(* Logix 5000 project; controller DSFW_0512_C_FCB_S1_SPN vendor 1 type 14 code 77 rev 20.12; software revision 20.06; part 2 of 3 *)
(* tags used below, declared in another part *)
   Alarms : DINT[3];
   Batch_Mode_Enable : BOOL;
   Comp_Low_Pressure_Alarm_Setpoint : REAL;
   Compressor_High_Pressure_Alarm_Setpoint : REAL;
   Compressor_High_Pressure_Delay_Timer : TIMER;
   Compressor_High_Superheat_Alarm_Delay : TIMER;
   Compressor_High_Superheat_Alarm_Setpoint : REAL;
   Compressor_Low_Pressure_Delay_Timer : TIMER;
   Compressor_Low_Subcooling_Alarm_Delay : TIMER;
   Compressor_Low_Subcooling_Alarm_Setpoint : REAL;
   Compressor_Low_Superheat_Alarm_Delay : TIMER;
   Compressor_Low_Superheat_Alarm_Setpoint : REAL;
   Compressor_OK_To_Run : BOOL;
   Compressor_Run_Proof_Delay : TIMER;
   Compressor_Short_Cycle_Time_Remaining : REAL;
   Compressor_Short_Cycle_Timer : TIMER;
   Compressor_Start_Delay : TIMER;
   Compressor_Subcooling : REAL;
   Compressor_Superheat : REAL;
   DV_IN_N7_100_199 : INT[10];
   DV_OUT_N7_0_99 : INT[20];
   EEV_101_Pressure_PIDE : PID_ENHANCED;
   EEV_101_Range_1_Max : REAL;
   EEV_101_Range_1_Min : REAL;
   EEV_101_Range_2_Max : REAL;
   EEV_101_Range_2_Min : REAL;
   EEV_101_Range_3_Max : REAL;
   EEV_101_Range_3_Min : REAL;
   EEV_101_Run_PIDE : BOOL;
   EEV_101_Run_Temp_PIDE : BOOL;
   EEV_101_Stop_PIDE : BOOL;
   EEV_101_Superheat_PIDE : PID_ENHANCED;
   EEV_101_Temperature_PIDE : PID_ENHANCED;
   EEV_102_Stop_PIDE : BOOL;
   Enable_Batch : BOOL;
   Evaporator_Superheat : REAL;
   Heaters_OK_To_Run : BOOL;
   Large_Batch_Derivative : REAL;
   Large_Batch_Integral : REAL;
   Large_Batch_Proportional : REAL;
   Large_Batch_Selected : BOOL;
   Medium_Batch_Derivative : REAL;
   Medium_Batch_Integral : REAL;
   Medium_Batch_Proportional : REAL;
   Medium_Batch_Selected : BOOL;
   PT_101_Offset : REAL;
   PT_101_Reactor_Supply_Pressure : REAL;
   PT_102_Compressor_Suction_Pressure : REAL;
   PT_102_Sensor_Alarm_Delay : TIMER;
   PT_103_Compressor_Discharge_Pressure : REAL;
   PT_103_Sensor_Alarm_Delay : TIMER;
   PT_104_Evaporator_Suction_Pressure : REAL;
   PT_104_Sensor_Alarm_Delay : TIMER;
   PT_105_Offset : REAL;
   PT_105_Tank_Blanket_Pressure : REAL;
   Pump_OK_To_Run : BOOL;
   Reaactor_Batch_PIDE : PID_ENHANCED;
   Reactor_Batch_CV_as_SP : REAL;
   Reactor_Batch_PID_Start : BOOL;
   Reactor_Batch_PID_Start_Delay : TIMER;
   Reactor_Batch_PID_Start_ONS : BOOL;
   Reactor_Batch_PID_Stop : BOOL;
   Reactor_Batch_PV : REAL;
   Reactor_Batch_SP_High : REAL;
   Reactor_Batch_SP_Low : REAL;
   Remote_Enable : BOOL;
   Remote_Start : BOOL;
   SCR_101_Auto_Manual : BOOL;
   SCR_101_Manual_Output : REAL;
   SCR_101_Run_PIDE : BOOL;
   SCR_101_Stop_PIDE : BOOL;
   SIC_101_Auto_Manual : BOOL;
   SIC_101_Manual_Output : REAL;
   SIC_101_Pressure_Setpoint : REAL;
   SIC_101_Run_PIDE : BOOL;
   SIC_101_Stop_PIDE : BOOL;
   Small_Batch_Derivative : REAL;
   Small_Batch_Integral : REAL;
   Small_Batch_Proportional : REAL;
   Small_Batch_Selected : BOOL;
   SP_Add_Max : REAL;
   System_Start : BOOL;
   TCV_101_Define_Range_1_Max : REAL;
   TCV_101_Define_Range_1_Min : REAL;
   TCV_101_Define_Range_2_Max : REAL;
   TCV_101_Define_Range_2_Min : REAL;
   TCV_101_Define_Range_3_Max : REAL;
   TCV_101_Define_Range_3_Min : REAL;
   TCV_101_PIDE : PID_ENHANCED;
   TCV_101_Range_1_Max : REAL;
   TCV_101_Range_1_Min : REAL;
   TCV_101_Range_2_Max : REAL;
   TCV_101_Range_2_Min : REAL;
   TCV_101_Range_3_Max : REAL;
   TCV_101_Range_3_Min : REAL;
   TCV_101_Run_PIDE : BOOL;
   TCV_101_Stop_PIDE : BOOL;
   TE_101_Liquid_Line_Temperature : REAL;
   TE_102_Evaporator_Suction_Temperature : REAL;
   TE_103_Compressor_Suction_Temperature : REAL;
   TE_104_Offset : REAL;
   TE_104_Reactor_Return_Temperature : REAL;
   TE_105_Offset : REAL;
   TE_105_Reactor_Supply_Temperature : REAL;
   Temperature_Setpoint : REAL;
   Test_Bit : BOOL[32];
   TIT_101_Offset : REAL;
   TIT_101_Vessel_Temperature : REAL;
   TIT_201_Vessel_Temperature : REAL;
   TIT_301_Vessel_Temperature : REAL;
   Vessel_1_Scale_Max : REAL;
   Vessel_1_Scale_Min : REAL;
   Vessel_1_Selected : BOOL;
   Vessel_2_Scale_Max : REAL;
   Vessel_2_Scale_Min : REAL;
   Vessel_2_Selected : BOOL;
   Vessel_3_Scale_Max : REAL;
   Vessel_3_Scale_Min : REAL;
   Vessel_3_Selected : BOOL;
(* Process_Control, continued *)

ROUTINE Heaters_Batch_Control   (* ladder *)
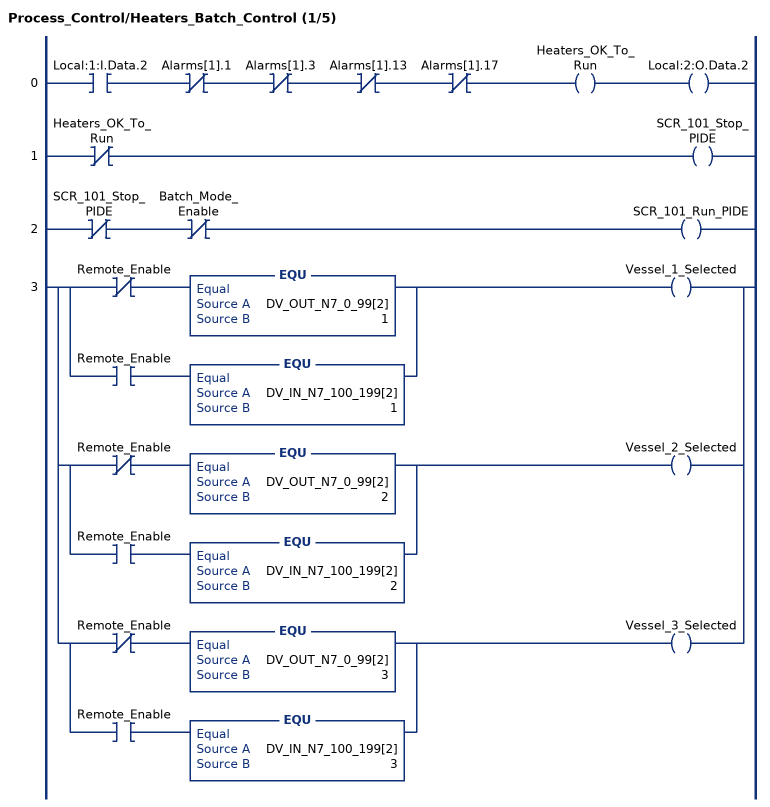
   0: XIC(Local:1:I.Data.2)XIO(Alarms[1].1)XIO(Alarms[1].3)XIO(Alarms[1].13)XIO(Alarms[1].17)OTE(Heaters_OK_To_Run)OTE(Local:2:O.Data.2);
   1: XIO(Heaters_OK_To_Run)OTE(SCR_101_Stop_PIDE);
   2: XIO(SCR_101_Stop_PIDE)XIO(Batch_Mode_Enable)OTE(SCR_101_Run_PIDE);
   3: [[XIO(Remote_Enable) EQU(DV_OUT_N7_0_99[2],1) ,XIC(Remote_Enable) EQU(DV_IN_N7_100_199[2],1) ] OTE(Vessel_1_Selected) ,[XIO(Remote_Enable) EQU(DV_OUT_N7_0_99[2],2) ,XIC(Remote_Enable) EQU(DV_IN_N7_100_199[2],2) ] OTE(Vessel_2_Selected) ,[XIO(Remote_Enable) EQU(DV_OUT_N7_0_99[2],3) ,XIC(Remote_Enable) EQU(DV_IN_N7_100_199[2],3) ] OTE(Vessel_3_Selected) ];
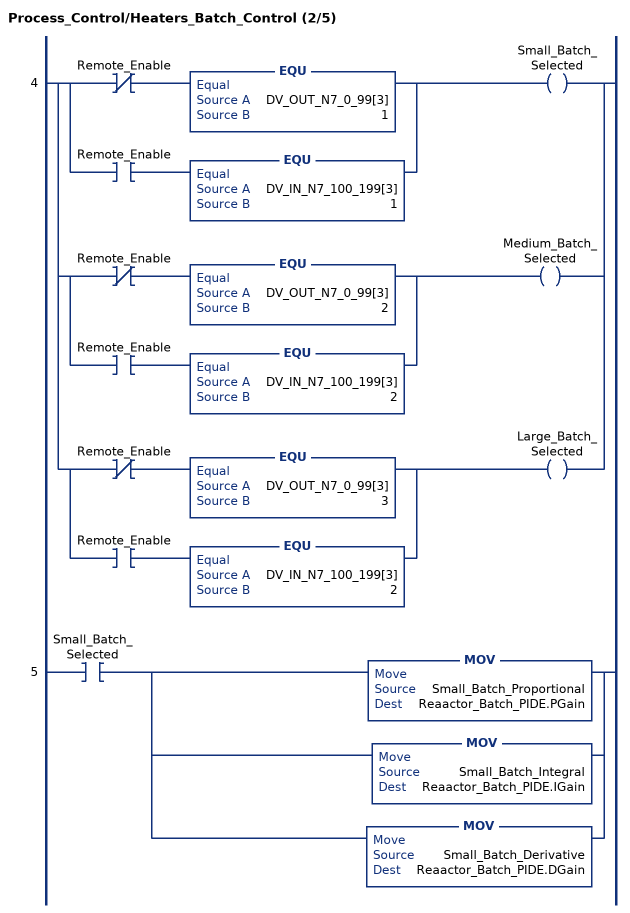
   4: [[XIO(Remote_Enable) EQU(DV_OUT_N7_0_99[3],1) ,XIC(Remote_Enable) EQU(DV_IN_N7_100_199[3],1) ] OTE(Small_Batch_Selected) ,[XIO(Remote_Enable) EQU(DV_OUT_N7_0_99[3],2) ,XIC(Remote_Enable) EQU(DV_IN_N7_100_199[3],2) ] OTE(Medium_Batch_Selected) ,[XIO(Remote_Enable) EQU(DV_OUT_N7_0_99[3],3) ,XIC(Remote_Enable) EQU(DV_IN_N7_100_199[3],2) ] OTE(Large_Batch_Selected) ];
   5: XIC(Small_Batch_Selected)[MOV(Small_Batch_Proportional,Reaactor_Batch_PIDE.PGain) ,MOV(Small_Batch_Integral,Reaactor_Batch_PIDE.IGain) ,MOV(Small_Batch_Derivative,Reaactor_Batch_PIDE.DGain) ];
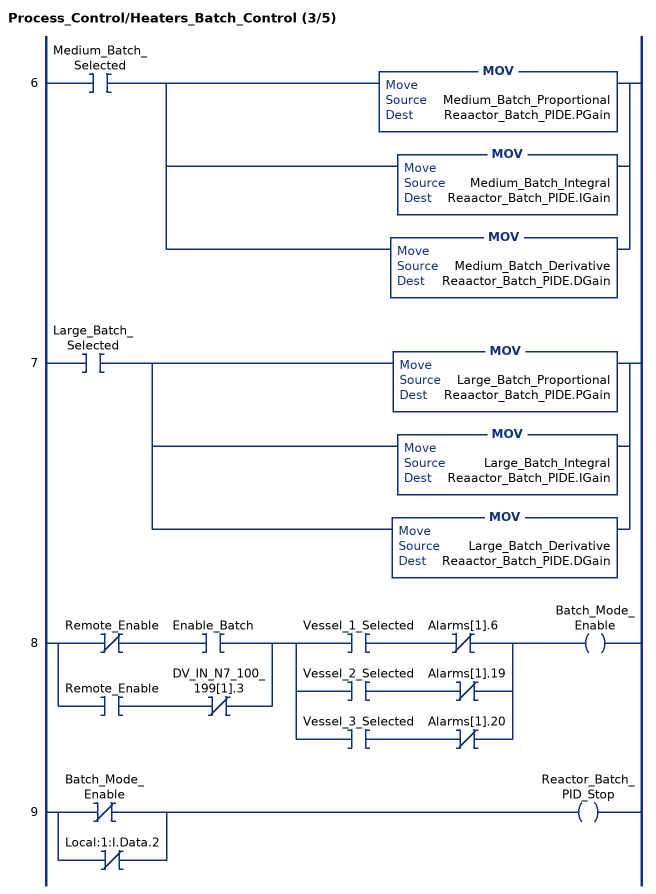
   6: XIC(Medium_Batch_Selected)[MOV(Medium_Batch_Proportional,Reaactor_Batch_PIDE.PGain) ,MOV(Medium_Batch_Integral,Reaactor_Batch_PIDE.IGain) ,MOV(Medium_Batch_Derivative,Reaactor_Batch_PIDE.DGain) ];
   7: XIC(Large_Batch_Selected)[MOV(Large_Batch_Proportional,Reaactor_Batch_PIDE.PGain) ,MOV(Large_Batch_Integral,Reaactor_Batch_PIDE.IGain) ,MOV(Large_Batch_Derivative,Reaactor_Batch_PIDE.DGain) ];
   8: [XIO(Remote_Enable) XIC(Enable_Batch) ,XIC(Remote_Enable) XIO(DV_IN_N7_100_199[1].3) ][XIC(Vessel_1_Selected) XIO(Alarms[1].6) ,XIC(Vessel_2_Selected) XIO(Alarms[1].19) ,XIC(Vessel_3_Selected) XIO(Alarms[1].20) ]OTE(Batch_Mode_Enable);
   9: [XIO(Batch_Mode_Enable) ,XIO(Local:1:I.Data.2) ]OTE(Reactor_Batch_PID_Stop);
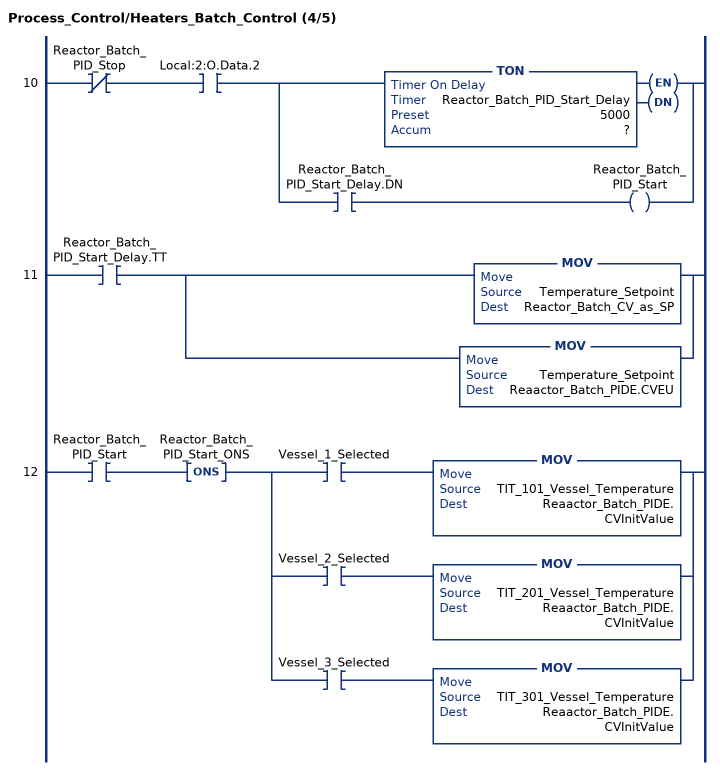
   10: XIO(Reactor_Batch_PID_Stop)XIC(Local:2:O.Data.2)[TON(Reactor_Batch_PID_Start_Delay,?,?) ,XIC(Reactor_Batch_PID_Start_Delay.DN) OTE(Reactor_Batch_PID_Start) ];
   11: XIC(Reactor_Batch_PID_Start_Delay.TT)[MOV(Temperature_Setpoint,Reactor_Batch_CV_as_SP) ,MOV(Temperature_Setpoint,Reaactor_Batch_PIDE.CVEU) ];
   12: XIC(Reactor_Batch_PID_Start)ONS(Reactor_Batch_PID_Start_ONS)[XIC(Vessel_1_Selected) MOV(TIT_101_Vessel_Temperature,Reaactor_Batch_PIDE.CVInitValue) ,XIC(Vessel_2_Selected) MOV(TIT_201_Vessel_Temperature,Reaactor_Batch_PIDE.CVInitValue) ,XIC(Vessel_3_Selected) MOV(TIT_301_Vessel_Temperature,Reaactor_Batch_PIDE.CVInitValue) ];
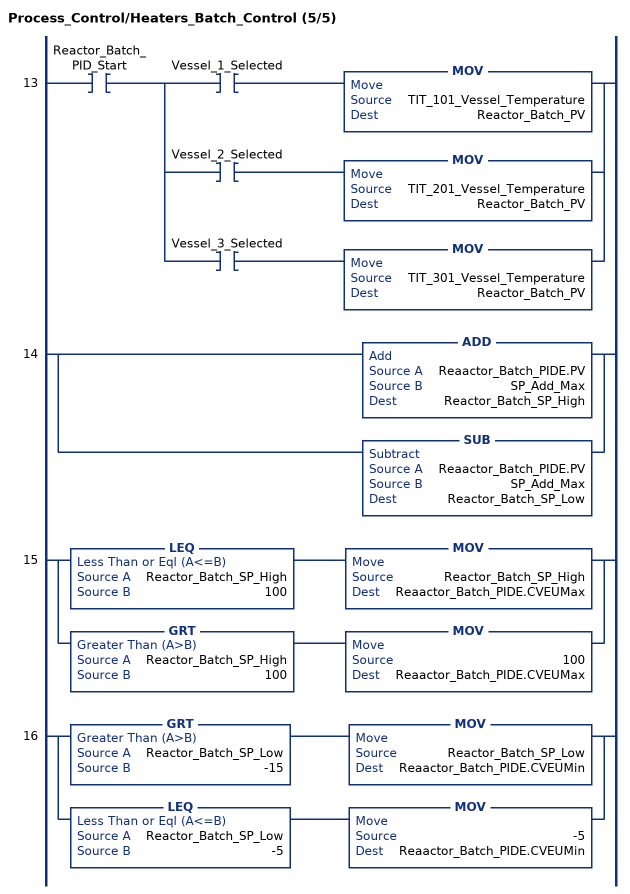
   13: XIC(Reactor_Batch_PID_Start)[XIC(Vessel_1_Selected) MOV(TIT_101_Vessel_Temperature,Reactor_Batch_PV) ,XIC(Vessel_2_Selected) MOV(TIT_201_Vessel_Temperature,Reactor_Batch_PV) ,XIC(Vessel_3_Selected) MOV(TIT_301_Vessel_Temperature,Reactor_Batch_PV) ];
   14: [ADD(Reaactor_Batch_PIDE.PV,SP_Add_Max,Reactor_Batch_SP_High) ,SUB(Reaactor_Batch_PIDE.PV,SP_Add_Max,Reactor_Batch_SP_Low) ];
   15: [LEQ(Reactor_Batch_SP_High,100) MOV(Reactor_Batch_SP_High,Reaactor_Batch_PIDE.CVEUMax) ,GRT(Reactor_Batch_SP_High,100) MOV(100,Reaactor_Batch_PIDE.CVEUMax) ];
   16: [GRT(Reactor_Batch_SP_Low,-15) MOV(Reactor_Batch_SP_Low,Reaactor_Batch_PIDE.CVEUMin) ,LEQ(Reactor_Batch_SP_Low,-5) MOV(-5,Reaactor_Batch_PIDE.CVEUMin) ];
END_ROUTINE

ROUTINE Pumps_Control   (* ladder *)
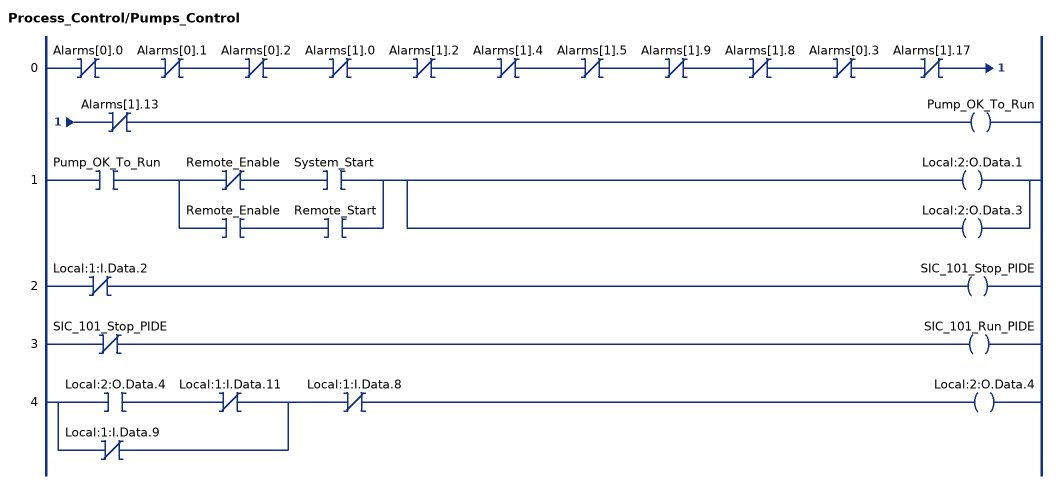
   0: XIO(Alarms[0].0)XIO(Alarms[0].1)XIO(Alarms[0].2)XIO(Alarms[1].0)XIO(Alarms[1].2)XIO(Alarms[1].4)XIO(Alarms[1].5)XIO(Alarms[1].9)XIO(Alarms[1].8)XIO(Alarms[0].3)XIO(Alarms[1].17)XIO(Alarms[1].13)OTE(Pump_OK_To_Run);
   1: XIC(Pump_OK_To_Run)[XIO(Remote_Enable) XIC(System_Start) ,XIC(Remote_Enable) XIC(Remote_Start) ][OTE(Local:2:O.Data.1) ,OTE(Local:2:O.Data.3) ];
   2: XIO(Local:1:I.Data.2)OTE(SIC_101_Stop_PIDE);
   3: XIO(SIC_101_Stop_PIDE)OTE(SIC_101_Run_PIDE);
   4: [XIC(Local:2:O.Data.4) XIO(Local:1:I.Data.11) ,XIO(Local:1:I.Data.9) ]XIO(Local:1:I.Data.8)OTE(Local:2:O.Data.4);
END_ROUTINE

ROUTINE Sensors   (* ladder *)
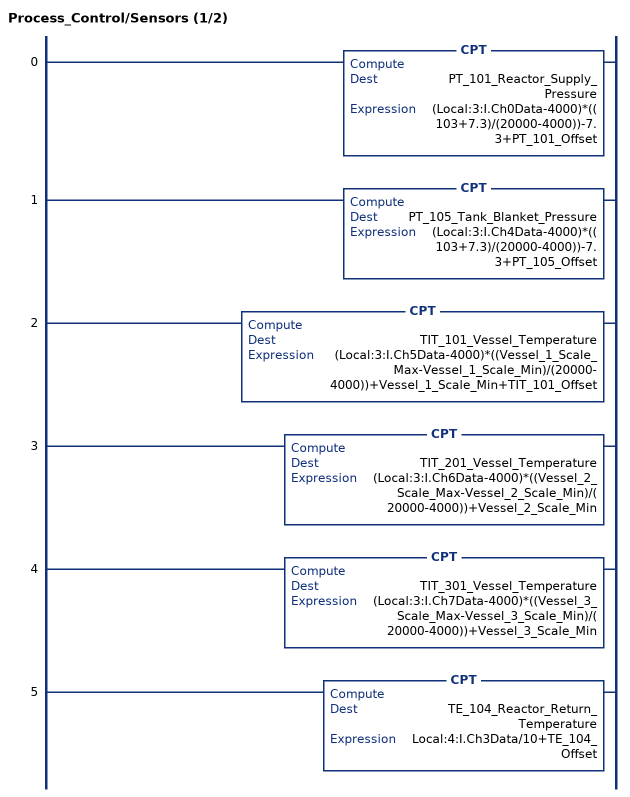
   0: CPT(PT_101_Reactor_Supply_Pressure,(Local:3:I.Ch0Data-4000)*((103+7.3)/(20000-4000))-7.3+PT_101_Offset);
   1: CPT(PT_105_Tank_Blanket_Pressure,(Local:3:I.Ch4Data-4000)*((103+7.3)/(20000-4000))-7.3+PT_105_Offset);
   2: CPT(TIT_101_Vessel_Temperature,(Local:3:I.Ch5Data-4000)*((Vessel_1_Scale_Max-Vessel_1_Scale_Min)/(20000-4000))+Vessel_1_Scale_Min+TIT_101_Offset);
   3: CPT(TIT_201_Vessel_Temperature,(Local:3:I.Ch6Data-4000)*((Vessel_2_Scale_Max-Vessel_2_Scale_Min)/(20000-4000))+Vessel_2_Scale_Min);
   4: CPT(TIT_301_Vessel_Temperature,(Local:3:I.Ch7Data-4000)*((Vessel_3_Scale_Max-Vessel_3_Scale_Min)/(20000-4000))+Vessel_3_Scale_Min);
   5: CPT(TE_104_Reactor_Return_Temperature,Local:4:I.Ch3Data/10+TE_104_Offset);
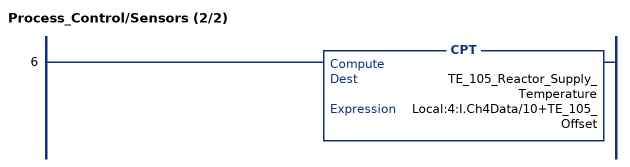
   6: CPT(TE_105_Reactor_Supply_Temperature,Local:4:I.Ch4Data/10+TE_105_Offset);
END_ROUTINE
END_PROGRAM

PROGRAM Process_PID_Calculations   (* main routine SIC_101 *)
VAR
   BOR_01 : FBD_BOOLEAN_OR := (In2 := 1, Out := 1);
   PIDE_01 : PID_ENHANCED := (PV := 40.73446, PVEUMax := 100.0, SPProg := 12.0, SPOper := 12.0, SPHLimit := 100.0, RatioProg := 1.0, RatioOper := 1.0, RatioHLimit := 1.0, RatioLLimit := 1.0, CVProg := 43.558277, CVOper := 43.558277, CVEUMax := 20000.0, CVEUMin := 4000.0, CVHLimit := 100.0, CVLLimit := 8.0, ControlAction := 1, PGain := 9.0, IGain := 1.9, PVEDerivative := 1, DSmoothing := 1, PVHHLimit := 150.0, PVHLimit := 100.0, PVLLimit := 2.0, PVLLLimit := 1.0, ProgValueReset := 1, RTSTime := 1, CVEU := 10969.324, CV := 43.558277, SP := 12.0, SPPercent := 12.0, PVPercent := 40.73446, E := 28.734459, EPercent := 28.734459, InitPrimary := 1, Ratio := 1.0, Auto := 1, DeltaT := 0.2);
   PIDE_02 : PID_ENHANCED := (PV := 40.73446, PVEUMax := 100.0, SPProg := 12.0, SPOper := 12.0, SPHLimit := 100.0, RatioProg := 1.0, RatioOper := 1.0, RatioHLimit := 1.0, RatioLLimit := 1.0, CVProg := 43.558277, CVOper := 43.558277, CVEUMax := 20000.0, CVEUMin := 4000.0, CVHLimit := 100.0, CVLLimit := 8.0, ControlAction := 1, PGain := 9.0, IGain := 1.9, PVEDerivative := 1, DSmoothing := 1, PVHHLimit := 150.0, PVHLimit := 100.0, PVLLimit := 2.0, PVLLLimit := 1.0, ProgValueReset := 1, RTSTime := 1, CVEU := 10969.324, CV := 43.558277, SP := 12.0, SPPercent := 12.0, PVPercent := 40.73446, E := 28.734459, EPercent := 28.734459, InitPrimary := 1, Ratio := 1.0, Auto := 1, DeltaT := 0.2);
END_VAR

ROUTINE SCR_101   (* function block diagram *)
   SHEET 1
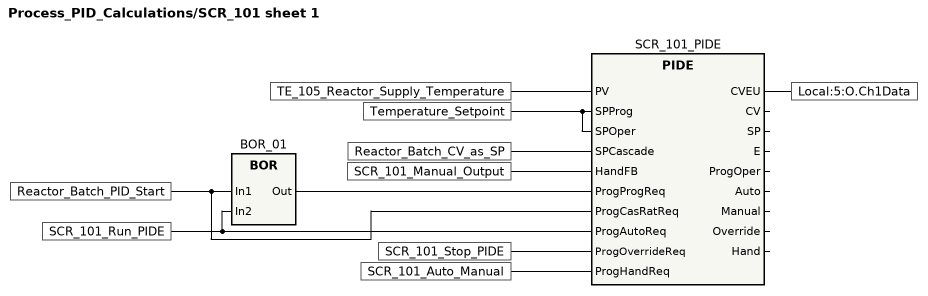
   BOR_01 : BOR(In1 := Reactor_Batch_PID_Start, In2 := SCR_101_Run_PIDE);
   SCR_101_PIDE : PIDE(PV := TE_105_Reactor_Supply_Temperature, SPProg := Temperature_Setpoint, SPOper := Temperature_Setpoint, SPCascade := Reactor_Batch_CV_as_SP, HandFB := SCR_101_Manual_Output, ProgProgReq := BOR_01.Out, ProgCasRatReq := Reactor_Batch_PID_Start, ProgAutoReq := SCR_101_Run_PIDE, ProgOverrideReq := SCR_101_Stop_PIDE, ProgHandReq := SCR_101_Auto_Manual);   // unwired pins: CV SP E ProgOper Auto Manual Override Hand
   Local:5:O.Ch1Data := SCR_101_PIDE.CVEU;
END_ROUTINE

ROUTINE SIC_101   (* function block diagram *)
   SHEET 1
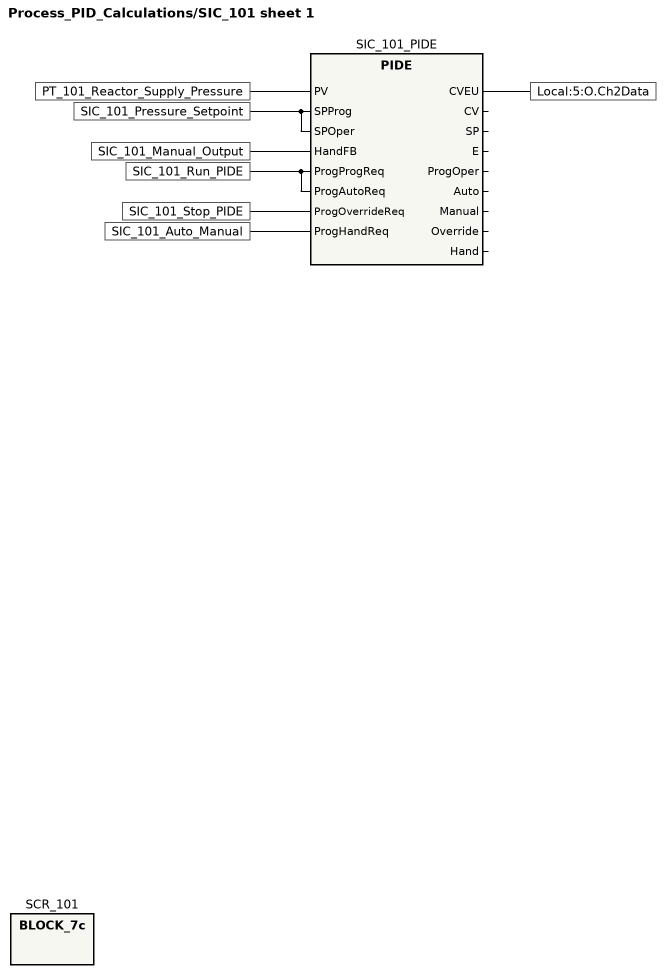
   SCR_101 : BLOCK_7c();
   SIC_101_PIDE : PIDE(PV := PT_101_Reactor_Supply_Pressure, SPProg := SIC_101_Pressure_Setpoint, SPOper := SIC_101_Pressure_Setpoint, HandFB := SIC_101_Manual_Output, ProgProgReq := SIC_101_Run_PIDE, ProgAutoReq := SIC_101_Run_PIDE, ProgOverrideReq := SIC_101_Stop_PIDE, ProgHandReq := SIC_101_Auto_Manual);   // unwired pins: CV SP E ProgOper Auto Manual Override Hand
   Local:5:O.Ch2Data := SIC_101_PIDE.CVEU;
END_ROUTINE
END_PROGRAM

PROGRAM Refrigeration_Control   (* main routine Config *)

ROUTINE Alarms   (* ladder *)
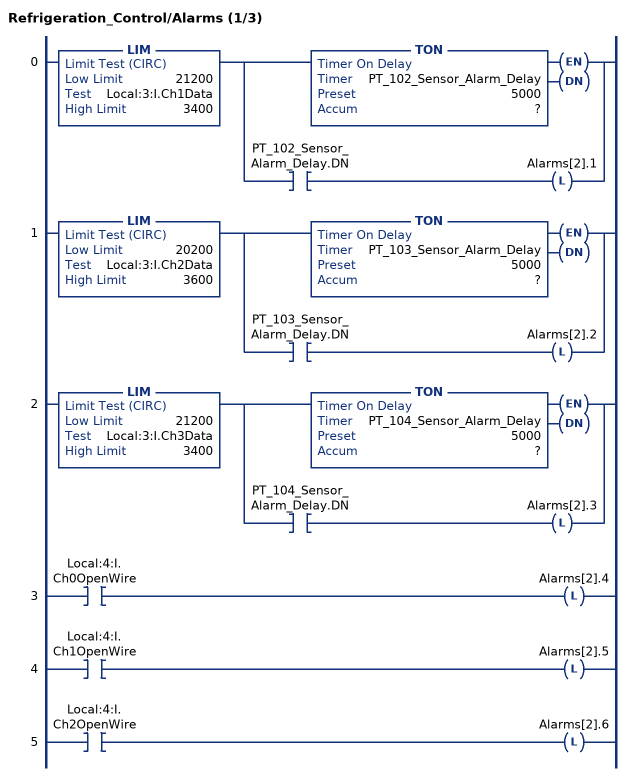
   0: LIM(21200,Local:3:I.Ch1Data,3400)[TON(PT_102_Sensor_Alarm_Delay,?,?) ,XIC(PT_102_Sensor_Alarm_Delay.DN) OTL(Alarms[2].1) ];
   1: LIM(20200,Local:3:I.Ch2Data,3600)[TON(PT_103_Sensor_Alarm_Delay,?,?) ,XIC(PT_103_Sensor_Alarm_Delay.DN) OTL(Alarms[2].2) ];
   2: LIM(21200,Local:3:I.Ch3Data,3400)[TON(PT_104_Sensor_Alarm_Delay,?,?) ,XIC(PT_104_Sensor_Alarm_Delay.DN) OTL(Alarms[2].3) ];
   3: XIC(Local:4:I.Ch0OpenWire)OTL(Alarms[2].4);
   4: XIC(Local:4:I.Ch1OpenWire)OTL(Alarms[2].5);
   5: XIC(Local:4:I.Ch2OpenWire)OTL(Alarms[2].6);
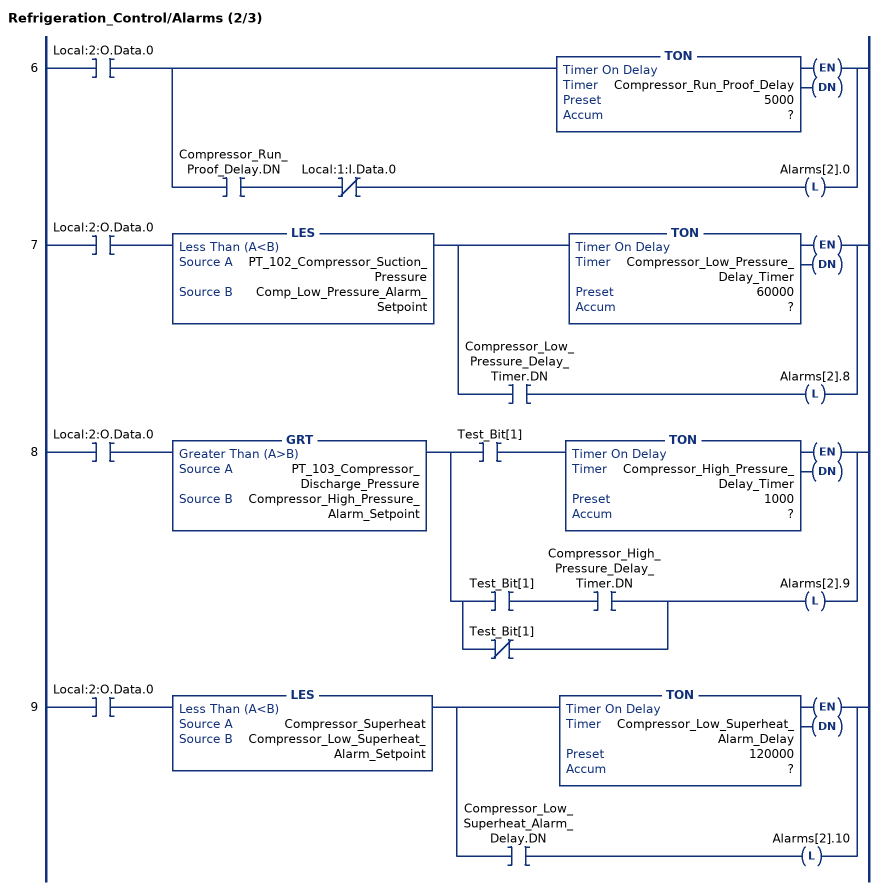
   6: XIC(Local:2:O.Data.0)[TON(Compressor_Run_Proof_Delay,?,?) ,XIC(Compressor_Run_Proof_Delay.DN) XIO(Local:1:I.Data.0) OTL(Alarms[2].0) ];
   7: XIC(Local:2:O.Data.0)LES(PT_102_Compressor_Suction_Pressure,Comp_Low_Pressure_Alarm_Setpoint)[TON(Compressor_Low_Pressure_Delay_Timer,?,?) ,XIC(Compressor_Low_Pressure_Delay_Timer.DN) OTL(Alarms[2].8) ];
   8: XIC(Local:2:O.Data.0)GRT(PT_103_Compressor_Discharge_Pressure,Compressor_High_Pressure_Alarm_Setpoint)[XIC(Test_Bit[1]) TON(Compressor_High_Pressure_Delay_Timer,?,?) ,[XIC(Test_Bit[1]) XIC(Compressor_High_Pressure_Delay_Timer.DN) ,XIO(Test_Bit[1]) ] OTL(Alarms[2].9) ];
   9: XIC(Local:2:O.Data.0)LES(Compressor_Superheat,Compressor_Low_Superheat_Alarm_Setpoint)[TON(Compressor_Low_Superheat_Alarm_Delay,?,?) ,XIC(Compressor_Low_Superheat_Alarm_Delay.DN) OTL(Alarms[2].10) ];
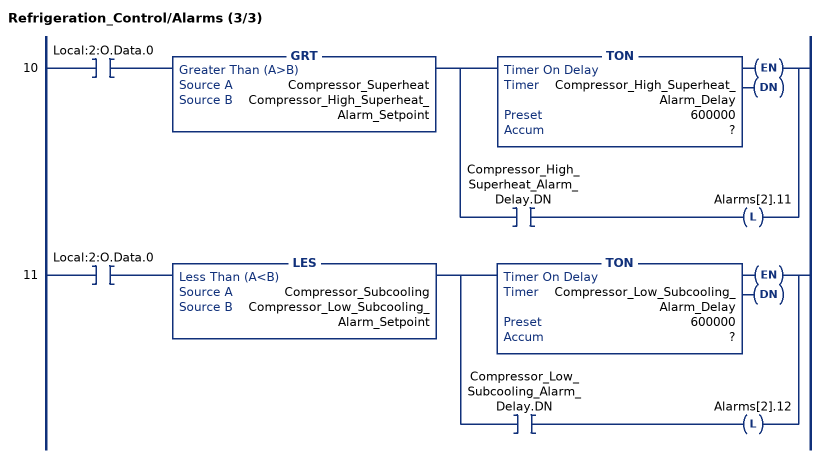
   10: XIC(Local:2:O.Data.0)GRT(Compressor_Superheat,Compressor_High_Superheat_Alarm_Setpoint)[TON(Compressor_High_Superheat_Alarm_Delay,?,?) ,XIC(Compressor_High_Superheat_Alarm_Delay.DN) OTL(Alarms[2].11) ];
   11: XIC(Local:2:O.Data.0)LES(Compressor_Subcooling,Compressor_Low_Subcooling_Alarm_Setpoint)[TON(Compressor_Low_Subcooling_Alarm_Delay,?,?) ,XIC(Compressor_Low_Subcooling_Alarm_Delay.DN) OTL(Alarms[2].12) ];
END_ROUTINE

ROUTINE Compressor_Control   (* ladder *)
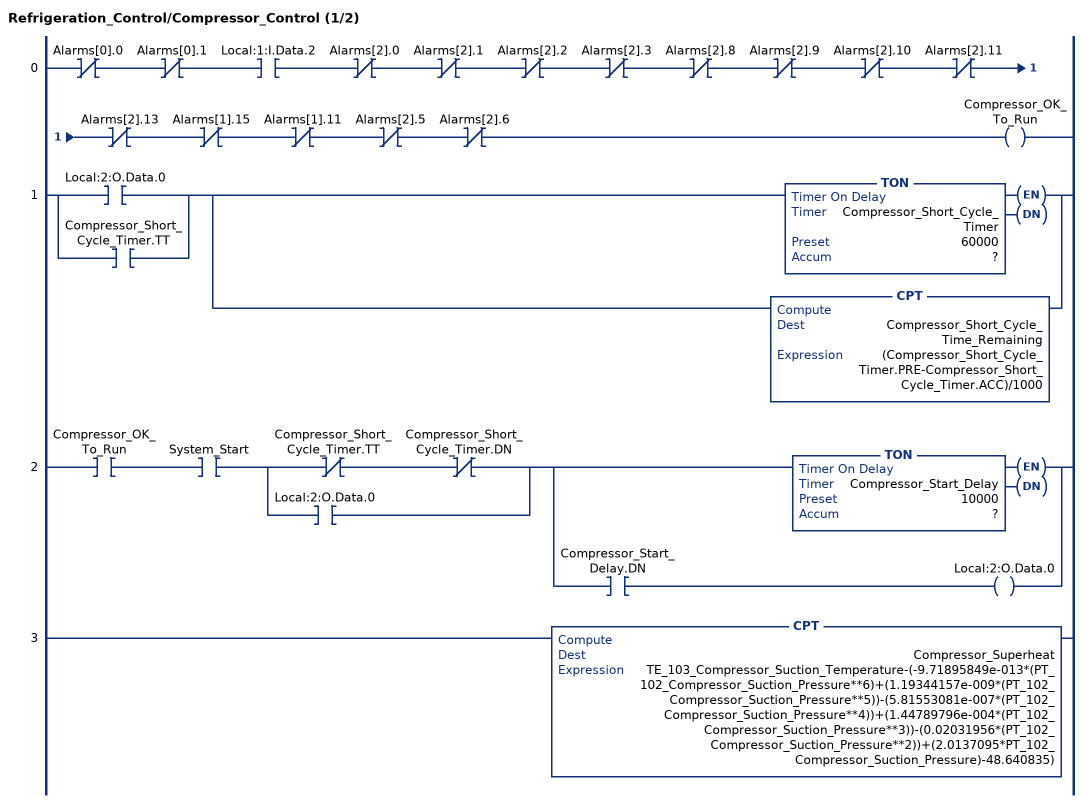
   0: XIO(Alarms[0].0)XIO(Alarms[0].1)XIC(Local:1:I.Data.2)XIO(Alarms[2].0)XIO(Alarms[2].1)XIO(Alarms[2].2)XIO(Alarms[2].3)XIO(Alarms[2].8)XIO(Alarms[2].9)XIO(Alarms[2].10)XIO(Alarms[2].11)XIO(Alarms[2].13)XIO(Alarms[1].15)XIO(Alarms[1].11)XIO(Alarms[2].5)XIO(Alarms[2].6)OTE(Compressor_OK_To_Run);
   1: [XIC(Local:2:O.Data.0) ,XIC(Compressor_Short_Cycle_Timer.TT) ][TON(Compressor_Short_Cycle_Timer,?,?) ,CPT(Compressor_Short_Cycle_Time_Remaining,(Compressor_Short_Cycle_Timer.PRE-Compressor_Short_Cycle_Timer.ACC)/1000) ];
   2: XIC(Compressor_OK_To_Run)XIC(System_Start)[XIO(Compressor_Short_Cycle_Timer.TT) XIO(Compressor_Short_Cycle_Timer.DN) ,XIC(Local:2:O.Data.0) ][TON(Compressor_Start_Delay,?,?) ,XIC(Compressor_Start_Delay.DN) OTE(Local:2:O.Data.0) ];
   3: CPT(Compressor_Superheat,TE_103_Compressor_Suction_Temperature-(-9.71895849e-013*(PT_102_Compressor_Suction_Pressure**6)+(1.19344157e-009*(PT_102_Compressor_Suction_Pressure**5))-(5.81553081e-007*(PT_102_Compressor_Suction_Pressure**4))+(1.44789796e-004*(PT_102_Compressor_Suction_Pressure**3))-(0.02031956*(PT_102_Compressor_Suction_Pressure**2))+(2.0137095*PT_102_Compressor_Suction_Pressure)-48.640835));
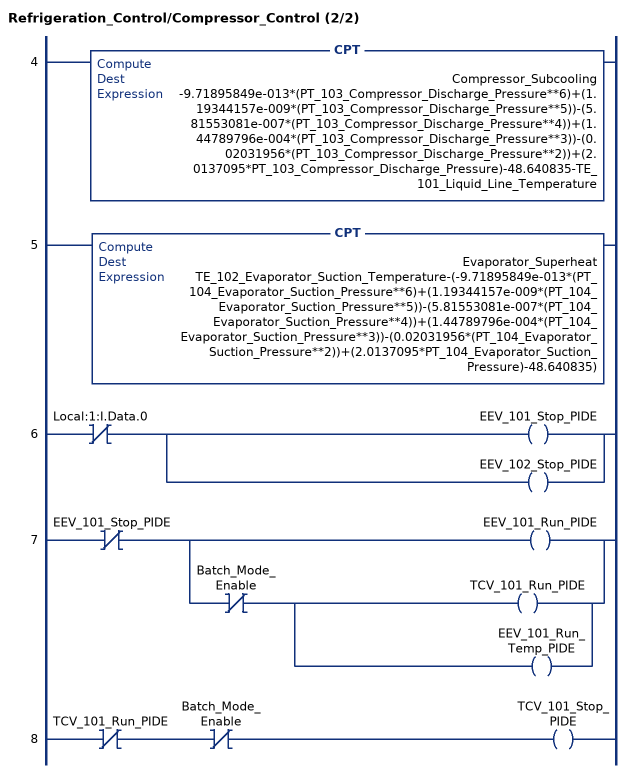
   4: CPT(Compressor_Subcooling,-9.71895849e-013*(PT_103_Compressor_Discharge_Pressure**6)+(1.19344157e-009*(PT_103_Compressor_Discharge_Pressure**5))-(5.81553081e-007*(PT_103_Compressor_Discharge_Pressure**4))+(1.44789796e-004*(PT_103_Compressor_Discharge_Pressure**3))-(0.02031956*(PT_103_Compressor_Discharge_Pressure**2))+(2.0137095*PT_103_Compressor_Discharge_Pressure)-48.640835-TE_101_Liquid_Line_Temperature);
   5: CPT(Evaporator_Superheat,TE_102_Evaporator_Suction_Temperature-(-9.71895849e-013*(PT_104_Evaporator_Suction_Pressure**6)+(1.19344157e-009*(PT_104_Evaporator_Suction_Pressure**5))-(5.81553081e-007*(PT_104_Evaporator_Suction_Pressure**4))+(1.44789796e-004*(PT_104_Evaporator_Suction_Pressure**3))-(0.02031956*(PT_104_Evaporator_Suction_Pressure**2))+(2.0137095*PT_104_Evaporator_Suction_Pressure)-48.640835));
   6: XIO(Local:1:I.Data.0)[OTE(EEV_101_Stop_PIDE) ,OTE(EEV_102_Stop_PIDE) ];
   7: XIO(EEV_101_Stop_PIDE)[OTE(EEV_101_Run_PIDE) ,XIO(Batch_Mode_Enable) [OTE(TCV_101_Run_PIDE) ,OTE(EEV_101_Run_Temp_PIDE) ] ];
   8: XIO(TCV_101_Run_PIDE)XIO(Batch_Mode_Enable)OTE(TCV_101_Stop_PIDE);
END_ROUTINE

ROUTINE Config   (* ladder *)
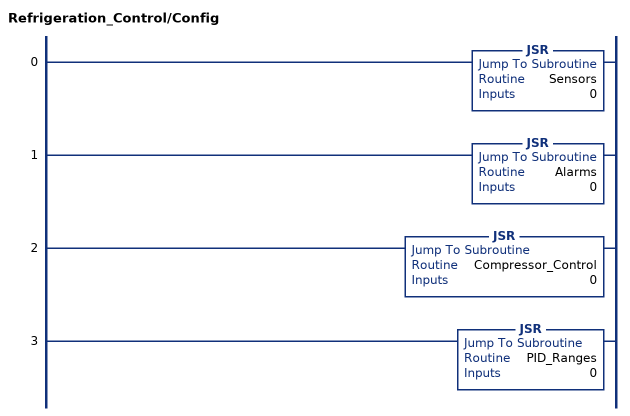
   0: JSR(Sensors,0);
   1: JSR(Alarms,0);
   2: JSR(Compressor_Control,0);
   3: JSR(PID_Ranges,0);
END_ROUTINE

ROUTINE PID_Ranges   (* ladder *)
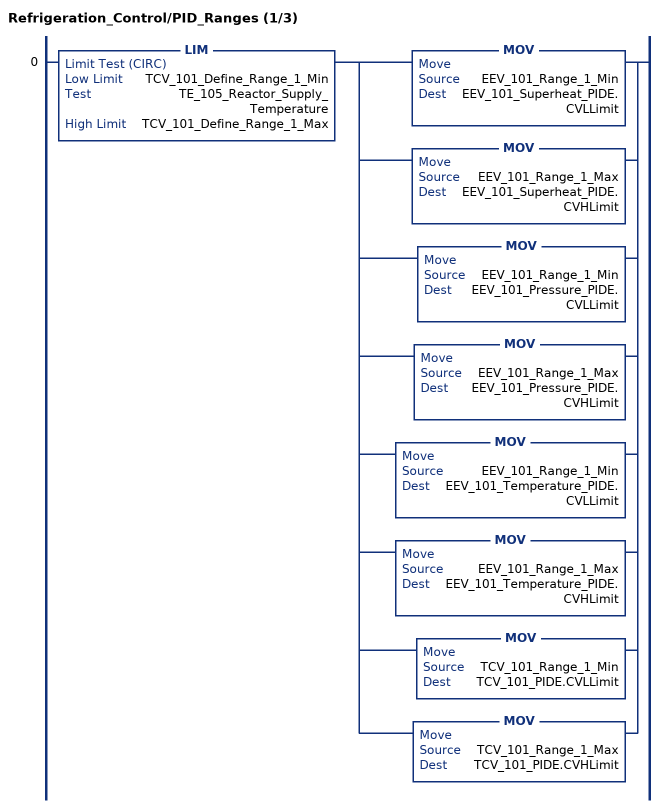
   0: LIM(TCV_101_Define_Range_1_Min,TE_105_Reactor_Supply_Temperature,TCV_101_Define_Range_1_Max)[MOV(EEV_101_Range_1_Min,EEV_101_Superheat_PIDE.CVLLimit) ,MOV(EEV_101_Range_1_Max,EEV_101_Superheat_PIDE.CVHLimit) ,MOV(EEV_101_Range_1_Min,EEV_101_Pressure_PIDE.CVLLimit) ,MOV(EEV_101_Range_1_Max,EEV_101_Pressure_PIDE.CVHLimit) ,MOV(EEV_101_Range_1_Min,EEV_101_Temperature_PIDE.CVLLimit) ,MOV(EEV_101_Range_1_Max,EEV_101_Temperature_PIDE.CVHLimit) ,MOV(TCV_101_Range_1_Min,TCV_101_PIDE.CVLLimit) ,MOV(TCV_101_Range_1_Max,TCV_101_PIDE.CVHLimit) ];
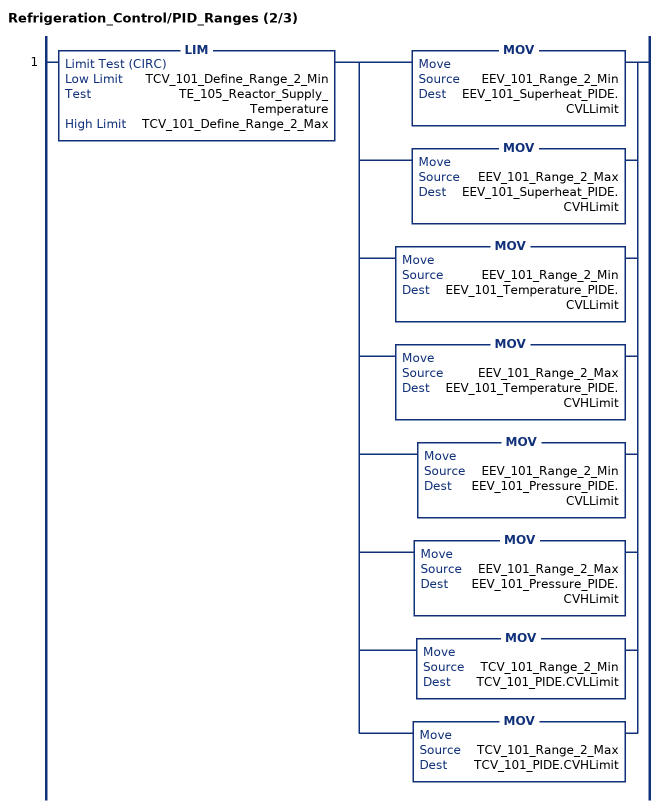
   1: LIM(TCV_101_Define_Range_2_Min,TE_105_Reactor_Supply_Temperature,TCV_101_Define_Range_2_Max)[MOV(EEV_101_Range_2_Min,EEV_101_Superheat_PIDE.CVLLimit) ,MOV(EEV_101_Range_2_Max,EEV_101_Superheat_PIDE.CVHLimit) ,MOV(EEV_101_Range_2_Min,EEV_101_Temperature_PIDE.CVLLimit) ,MOV(EEV_101_Range_2_Max,EEV_101_Temperature_PIDE.CVHLimit) ,MOV(EEV_101_Range_2_Min,EEV_101_Pressure_PIDE.CVLLimit) ,MOV(EEV_101_Range_2_Max,EEV_101_Pressure_PIDE.CVHLimit) ,MOV(TCV_101_Range_2_Min,TCV_101_PIDE.CVLLimit) ,MOV(TCV_101_Range_2_Max,TCV_101_PIDE.CVHLimit) ];
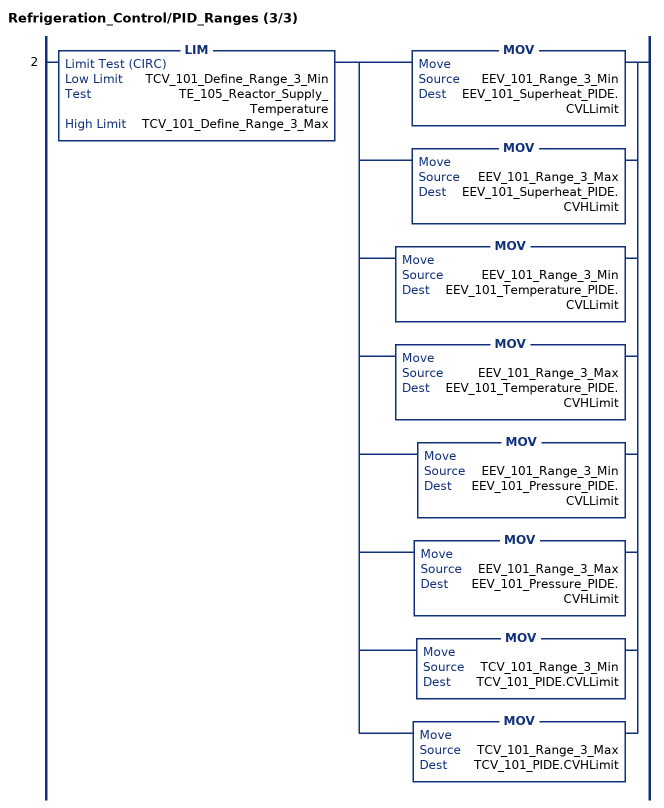
   2: LIM(TCV_101_Define_Range_3_Min,TE_105_Reactor_Supply_Temperature,TCV_101_Define_Range_3_Max)[MOV(EEV_101_Range_3_Min,EEV_101_Superheat_PIDE.CVLLimit) ,MOV(EEV_101_Range_3_Max,EEV_101_Superheat_PIDE.CVHLimit) ,MOV(EEV_101_Range_3_Min,EEV_101_Temperature_PIDE.CVLLimit) ,MOV(EEV_101_Range_3_Max,EEV_101_Temperature_PIDE.CVHLimit) ,MOV(EEV_101_Range_3_Min,EEV_101_Pressure_PIDE.CVLLimit) ,MOV(EEV_101_Range_3_Max,EEV_101_Pressure_PIDE.CVHLimit) ,MOV(TCV_101_Range_3_Min,TCV_101_PIDE.CVLLimit) ,MOV(TCV_101_Range_3_Max,TCV_101_PIDE.CVHLimit) ];
END_ROUTINE
